// TIA Portal V20 export
// export: Created 2026-10-12T04:58:23.0872973Z, ExportSetting WithDefaults, DisplayName Totally Integrated Automation Portal, DisplayVersion V20, DisplayName TIA Portal Openness, DisplayVersion V20, DisplayName TIA Portal Teamcenter Gateway, DisplayVersion V20, DisplayName TIA Portal Version Control Interface, DisplayVersion V20, DisplayName SINAMICS Startdrive Advanced, DisplayVersion V20 SP1 Update 2, DisplayName SINAMICS Startdrive G110M, G120, G120C, G120D, G120P, G115D, DisplayVersion V20 SP1 Update 2, DisplayName SINAMICS Startdrive G130, G150, S120, S150, SINAMICS MV, G220, S200, S210, DisplayVersion V20 SP1 Update 2, DisplayName STEP 7 Professional, DisplayVersion V20, DisplayName STEP 7 Safety, DisplayVersion V20, DisplayName WinCC Basic/Comfort/Advanced, DisplayVersion V20, DisplayName WinCC Professional, DisplayVersion V20, DisplayName WinCC Unified, DisplayVersion V20
FUNCTION "FRK_Config_DeclarationCell" : Void   // FC133, SCL
{ S7_Optimized_Access := 'TRUE' }
VERSION : 0.1
// stored: AutoNumber true, IsIECCheckEnabled false, SetENOAutomatically false, UDAEnableTagReadback false
   VAR_INPUT
      Access : "FRK_Access";
      RootIndex : Int;
      ModelIndex : UDInt;
   END_VAR
   VAR_IN_OUT
      Module : "FB_DeclarationCell";
      Cursor : "FRK_ConfigCursor";
      Page : "ST_ConfigPage";
   END_VAR
   VAR_TEMP
      Ok : Bool;
   END_VAR
BEGIN

   IF #ModelIndex = 0 THEN
       "FRK_ConfigCatalog"(Scope := #Module.Status.Name,
                           Catalog := #Module.Catalog,
                           Count := #Module.CatalogCount,
                           ReadLevel := #Access.Policy.Required[0],
                           Readable := #Access.CurrentLevel >= #Access.Policy.Required[0],
                           Cursor := #Cursor,
                           Page := #Page);
   END_IF;
   IF #ModelIndex = 0 THEN
       "FRK_CfgDef_DeclarationCell"(FieldIndex := 1);
       "FRK_ConfigScratch".Entry.Scope := STRING_TO_WSTRING(#Module.Status.Name);
       "FRK_ConfigScratch".Entry.ReadLevel := MAX(IN1 := #Access.Policy.Required[0], IN2 := "FRK_ConfigScratch".MinRead);
       "FRK_ConfigScratch".Entry.WriteLevel := MAX(IN1 := #Access.Policy.Required[1], IN2 := "FRK_ConfigScratch".MinWrite);
       "FRK_ConfigScratch".Entry.Readable := #Access.CurrentLevel >= "FRK_ConfigScratch".Entry.ReadLevel;
       "FRK_ConfigScratch".Entry.ModelScoped := FALSE;
       "FRK_ConfigScratch".Entry.ValueText := DINT_TO_WSTRING(TIME_TO_DINT(#Module.ParCfg.Timeout));
       IF NOT "FRK_ConfigScratch".Entry.Readable THEN
           "FRK_ConfigScratch".Entry.ValueText := WSTRING#'';
       END_IF;
       "FRK_ConfigAppendEntry"(Cursor := #Cursor,
                               Page := #Page);
   END_IF;
   IF #ModelIndex = 0 THEN
       "FRK_CfgDef_DeclarationCell"(FieldIndex := 2);
       "FRK_ConfigScratch".Entry.Scope := STRING_TO_WSTRING(#Module.Status.Name);
       "FRK_ConfigScratch".Entry.ReadLevel := MAX(IN1 := #Access.Policy.Required[0], IN2 := "FRK_ConfigScratch".MinRead);
       "FRK_ConfigScratch".Entry.WriteLevel := MAX(IN1 := #Access.Policy.Required[1], IN2 := "FRK_ConfigScratch".MinWrite);
       "FRK_ConfigScratch".Entry.Readable := #Access.CurrentLevel >= "FRK_ConfigScratch".Entry.ReadLevel;
       "FRK_ConfigScratch".Entry.ModelScoped := FALSE;
       "FRK_ConfigScratch".Entry.ValueText := DINT_TO_WSTRING(#Module.ParCfg.Preset);
       IF NOT "FRK_ConfigScratch".Entry.Readable THEN
           "FRK_ConfigScratch".Entry.ValueText := WSTRING#'';
       END_IF;
       "FRK_ConfigAppendEntry"(Cursor := #Cursor,
                               Page := #Page);
   END_IF;
   IF #ModelIndex = 0 THEN
       "FRK_Config_DeclarationCylinder"(Module := #Module.Clamp,
                                        Access := #Access,
                                        RootIndex := #RootIndex,
                                        ModelIndex := #ModelIndex,
                                        Cursor := #Cursor,
                                        Page := #Page);
   END_IF;
   IF #ModelIndex = 0 THEN
       "FRK_Config_DeclarationCylinder"(Module := #Module.Gate,
                                        Access := #Access,
                                        RootIndex := #RootIndex,
                                        ModelIndex := #ModelIndex,
                                        Cursor := #Cursor,
                                        Page := #Page);
   END_IF;
END_FUNCTION
